(*
SPDX-FileCopyrightText: c 2026 Oleksandr Tiutyk <trofimich@gmail.com>
SPDX-License-Identifier: MIT
License: https://opensource.org/license/mit
*)

(*!
<summary>Checks ascending sorting of a full list with duplicate strings and reverse lookup.</summary>
<description>
Owns a list and its copied entries. Use from one task at a stable address.
Teardown clears surviving entries before publication.
</description>
*)

{attribute 'no_assign'}
{attribute 'no_explicit_call' := 'do not call this function block directly'}
FUNCTION_BLOCK StaticListSortTest EXTENDS TOF_Testing.SingleCycleTest
VAR_STAT
	{attribute 'hide'}
	_ClassName : STRING := __POUNAME();
END_VAR
VAR
	_List : TOF_Collections.List<8>(valueValidator := 0);
	_Predicate : ListStringPredicate;
END_VAR

(*!
<summary>Checks ascending sorting of a full list with duplicate strings and reverse lookup.</summary>
*)
METHOD PROTECTED ExecuteTest
VAR
	values : ARRAY [0..5] OF STRING := ['String0', 'String1', 'String2', 'String3', 'String4', 'String5'];
	expected : ARRAY [0..7] OF STRING :=
		['String0', 'String1', 'String2', 'String2', 'String2', 'String3', 'String4', 'String5'];
	i : DINT;
	index : TOF_Core.DINT_INDEX;
	found : BOOL;
	entry : TOF_Core.GENERIC_VALUE;
END_VAR
_List.AppendCopy(value := values[5]);
_List.AppendCopy(value := values[4]);
_List.AppendCopy(value := values[3]);
_List.AppendCopy(value := values[2]);
_List.AppendCopy(value := values[2]);
_List.AppendCopy(value := values[2]);
_List.AppendCopy(value := values[1]);
_List.AppendCopy(value := values[0]);

_List.Sort(comparer := TOF_Comparison.StandardComparers.StringComparer);

Assert.ThatDInt(
	actual := _List.Length,
	message := "Ascending sort length"
).ToBe(expected := DINT#8);

FOR i := 0 TO 7 DO
	Assert.ThatString(
		actual := _List.Get(index := i).AsString255(),
		message := TOF_Core.WideStrings.Concat255("Ascending sort at index ", TO_WSTRING(i))
	).ToBe(expected := expected[i]);
END_FOR

_Predicate.Expected := 'String3';

found := _List.FindSingle(
	predicate := _Predicate,
	searchDirection := TOF_Core.SEARCH_DIRECTION.FROM_END,
	value => entry,
	index => index
);

Assert.ThatBool(
	actual := found AND_THEN index = 5 AND_THEN entry.AsString255() = 'String3',
	message := "Reverse lookup must return String3 at its current position after sorting"
).IsTrue();
END_METHOD

(*!
<summary>Clears the fixture before the runner publishes the result.</summary>
<description>
Also runs after an unexpected exception interrupts the case.
</description>
*)
METHOD PROTECTED AfterTest
_List.Clear();
END_METHOD

//! <summary>Borrows the concrete class name. Callers must not modify it.</summary>
{attribute 'monitoring' := 'call'}
PROPERTY ClassName : REFERENCE TO STRING
GET
ClassName REF= _ClassName;
END_GET
END_PROPERTY

//! <summary>Borrows the compiler-initialized namespace name. Callers must not modify it.</summary>
{attribute 'monitoring' := 'call'}
PROPERTY NamespaceName : REFERENCE TO STRING
GET
NamespaceName REF= CurrentNamespace.Name;
END_GET
END_PROPERTY

//! <summary>Reports the concrete instance size in bytes.</summary>
{attribute 'monitoring' := 'call'}
PROPERTY SelfSize : ULINT
GET
SelfSize := XSIZEOF(THIS^);
END_GET
END_PROPERTY

END_FUNCTION_BLOCK

(* stored: Version 1.1.0.1
   POU StaticListSortTest: Id {51d42083-1ba6-41c3-9c5e-e61724ad606b}, SpecialFunc None
   Method ExecuteTest: Id {1b29d960-ae20-4bae-8d3d-5409e3ba5a8c}
   Method AfterTest: Id {1eb7a9d1-f4b3-4c3d-b61b-106ec1b25383}
   Property ClassName: Id {82572386-b38c-4430-9477-4e0e8169ea1a}
   Get Get: Id {3a5553e1-98c7-4021-91a0-5556ff11f2eb}
   Property NamespaceName: Id {db22e762-906e-4993-8c49-dae5a6eb888f}
   Get Get: Id {b07a5ebc-e5fc-4e4c-82e2-1684d158bd29}
   Property SelfSize: Id {6dbaf7ed-cdd7-461d-bafc-d258fe5c95d5}
   Get Get: Id {ae0952d9-ca12-4be2-8e06-73e8c4370a88} *)
